Fanuc KAREL source: kt00402.KL

-- PROVISIONAL review KL for V1013-1; original PC SHA256 e6514f2490f8e75bf44f248af42a69a91faa322880040e31e799a4ff35a41149
-- Incomplete behavior may be omitted. Consult companion uncertainty JSON. Do not deploy.
PROGRAM KT00402
%NOLOCKGROUP
VAR
  I1 : INTEGER
  R2 : REAL
  OUT : BOOLEAN
BEGIN
  -- UNRESOLVED_PC offsets 5-16; opcodes 2E,23
  -- UNRESOLVED_PC offsets 21-32; opcodes 2E,23
  -- UNRESOLVED_PC offsets 37-59; opcodes 21,21,29,64,29,71,23
  -- UNRESOLVED_PC offsets 64-68; opcodes 7F
END KT00402
